// TIA Portal V21 export
// export: Created 2026-11-08T21:17:29.1331056Z, ExportSetting WithDefaults, DisplayName Totally Integrated Automation Portal, DisplayVersion V21 Update 3, DisplayName STEP 7 Professional, DisplayVersion V21 Update 3, DisplayName STEP 7 Safety, DisplayVersion V21, DisplayName Tech WebApplication, DisplayVersion V21, DisplayName WinCC Basic/Comfort/Advanced, DisplayVersion V21 Update 3, DisplayName WinCC Unified, DisplayVersion V21 Update 3
DATA_BLOCK "DB_OfUdt"   // DB8
{ S7_Optimized_Access := 'TRUE' }
VERSION : 0.1
// stored: AutoNumber true, DBAccessibleFromOPCUA true, DBAccessibleFromWebserver true, InstanceOfName UDT_Outer, InstanceOfType UDT, IsOnlyStoredInLoadMemory false, IsWriteProtectedInAS false
"UDT_Outer"
   // VAR
   //    inner { S7_SetPoint := 'True'} : "UDT_Inner";
   //    innerArr { S7_SetPoint := 'True'} : Array[0..1] of "UDT_Inner";
   //    s : Struct
   //       "a" : Bool;
   //       "m" : Array[0..1, 0..1] of Byte;
   //    END_STRUCT;
   //    txt : String[20] := 'udtdb';
   // END_VAR
BEGIN
   inner.Temp := 1.0;
END_DATA_BLOCK
